(* IEC 61131-3 sources: kauha-loader-autonomy/plc/codesys/src, 6 files *)

(* ---- DUT_Types.st ---- *)
(* KAUHA safety PLC: data types.
   IEC 61131-3 Structured Text, 2nd edition subset (no methods, no references),
   so the same source compiles in CODESYS and in the matiec compiler the tests use. *)

TYPE ST_SafetyConfig :
STRUCT
    (* SafetyParams *)
    remote_timeout_s     : LREAL;
    watchdog_timeout_s   : LREAL;
    overspeed_tol        : LREAL;
    decel_ramp           : LREAL;
    ramp_reaction_s      : LREAL;
    discrepancy_tol      : LREAL;
    discrepancy_time_s   : LREAL;
    position_invalid_s   : LREAL;
    max_mute_s           : LREAL;
    auto_restart_clear_s : LREAL;
    warning_hold_s       : LREAL;
    auto_speed           : LREAL;
    teleop_speed         : LREAL;
    warning_speed        : LREAL;
    standstill           : LREAL;
    recovery_speed       : LREAL;
    side_recovery_speed  : LREAL;
    (* FieldTable: facts about the field sets loaded into the scanners *)
    t_standstill         : LREAL;
    dig_speed            : LREAL;
    dock_speed           : LREAL;
    speed_cap            : LREAL;
    auto_restart         : BOOL;     (* SR-11 automatic restart after a clearing stop *)
    band0                : LREAL;    (* speed band tops, m/s *)
    band1                : LREAL;
    band2                : LREAL;
    band3                : LREAL;
    sector0              : LREAL;    (* articulation sector boundaries, rad *)
    sector1              : LREAL;
    sector2              : LREAL;
    sector3              : LREAL;
    vprot0               : LREAL;    (* highest speed each band's protective field stops from *)
    vprot1               : LREAL;
    vprot2               : LREAL;
    vprot3               : LREAL;
    n_sectors            : INT;
    n_bands              : INT;
END_STRUCT;
END_TYPE

TYPE ST_SafetyInputs :
STRUCT
    t                : LREAL;   (* monotonic time, s *)
    mode             : INT;     (* 0 IDLE, 1 AUTO, 2 TELEOP *)
    speed_a          : LREAL;   (* drive-by-wire gateway, non-safety source, m/s *)
    speed_b          : LREAL;   (* PLC's own speed sensor, m/s *)
    articulation     : LREAL;   (* PLC's own articulation sensor, rad *)
    front_prot       : BOOL;
    front_warn       : BOOL;
    rear_prot        : BOOL;
    rear_warn        : BOOL;
    side_prot        : BOOL;
    side_contact     : BOOL;
    scanners_ok      : BOOL;
    remote_hb_age    : LREAL;
    remote_estop     : BOOL;
    reset_req        : BOOL;
    machine_estop    : BOOL;
    autonomy_cmd_age : LREAL;
    dig_req          : BOOL;
    dock_req         : BOOL;
    in_operating_area : BOOL;
    in_dig_zone      : BOOL;
    in_dock_zone     : BOOL;
    truck_door_open  : BOOL;
    boom_raised      : BOOL;
    front_side       : BOOL;
    under_near       : BOOL;
    under_far        : BOOL;
    under_mid        : BOOL;
    position_valid   : BOOL;
END_STRUCT;
END_TYPE

TYPE ST_SafetyOutputs :
STRUCT
    state            : INT;     (* 0 RUN, 1 WARNING, 2 PROTECTIVE_STOP, 3 EMERGENCY_STOP *)
    cause            : WORD;    (* latched causes, bit mask as in kauha/safety/core.py *)
    speed_limit      : LREAL;
    field_set        : INT;
    brake_release    : BOOL;    (* FALSE: drive power cut, motors short-braked (hardwired) *)
    implement_enable : BOOL;    (* FALSE: actuator power cut (hardwired) *)
    reset_pending    : BOOL;
    dock_blocked     : BOOL;
    fs_direction     : INT;
    fs_v_protected   : LREAL;
    recovery         : WORD;    (* fields in SR-12 recovery *)
    ev_stop          : BOOL;    (* a stop event was logged this cycle *)
    ev_recovery      : BOOL;
    ev_reset         : BOOL;
END_STRUCT;
END_TYPE

(* Eight payload bytes. A struct, not a bare array type, so it can be passed to
   functions by value in every IEC compiler (matiec mis-handles bare array types). *)
TYPE ST_Payload :
STRUCT
    b : ARRAY [0..7] OF BYTE;
END_STRUCT;
END_TYPE

TYPE ST_Frame :
STRUCT
    id   : DWORD;                    (* 29-bit J1939 identifier *)
    data : ST_Payload;
END_STRUCT;
END_TYPE

(* ---- GVL_Config.st ---- *)
(* KAUHA safety configuration lists, one per profile. Select one in PRG_Safety. *)

(* Generated by kauha.scale.profile for profile 'full'. Do not edit by hand. *)
VAR_GLOBAL CONSTANT
    CFG_FULL : ST_SafetyConfig := (
        remote_timeout_s := 0.5,
        watchdog_timeout_s := 0.2,
        overspeed_tol := 0.2,
        decel_ramp := 0.8,
        ramp_reaction_s := 0.3,
        discrepancy_tol := 0.3,
        discrepancy_time_s := 0.2,
        position_invalid_s := 2,
        max_mute_s := 25,
        auto_restart_clear_s := 3,
        warning_hold_s := 2,
        auto_speed := 3,
        teleop_speed := 3,
        warning_speed := 1,
        standstill := 0.05,
        recovery_speed := 0.5,
        side_recovery_speed := 0.3,
        t_standstill := 0.1,
        dig_speed := 1,
        dock_speed := 0.6,
        speed_cap := 2.97018412,
        auto_restart := TRUE,
        band0 := 0.5,
        band1 := 1.5,
        band2 := 2.5,
        band3 := 3,
        sector0 := -0.3,
        sector1 := -0.1,
        sector2 := 0.1,
        sector3 := 0.3,
        vprot0 := 0.794930202,
        vprot1 := 1.5,
        vprot2 := 2.5,
        vprot3 := 3.17018412,
        n_sectors := 5,
        n_bands := 4
    );
END_VAR

(* Generated by kauha.scale.profile for profile 'scale8_nanoscan3'. Do not edit by hand. *)
VAR_GLOBAL CONSTANT
    CFG_SCALE8_NANOSCAN3 : ST_SafetyConfig := (
        remote_timeout_s := 0.5,
        watchdog_timeout_s := 0.2,
        overspeed_tol := 0.0707106781,
        decel_ramp := 0.8,
        ramp_reaction_s := 0.1,
        discrepancy_tol := 0.106066017,
        discrepancy_time_s := 0.2,
        position_invalid_s := 2,
        max_mute_s := 8.83883476,
        auto_restart_clear_s := 1.06066017,
        warning_hold_s := 0.707106781,
        auto_speed := 1.06066017,
        teleop_speed := 1.06066017,
        warning_speed := 0.353553391,
        standstill := 0.0176776695,
        recovery_speed := 0.176776695,
        side_recovery_speed := 0.106066017,
        t_standstill := 0.0353553391,
        dig_speed := 0.353553391,
        dock_speed := 0.212132034,
        speed_cap := 1.00147274,
        auto_restart := TRUE,
        band0 := 0.176776695,
        band1 := 0.530330086,
        band2 := 0.883883476,
        band3 := 1.06066017,
        sector0 := -0.3,
        sector1 := -0.1,
        sector2 := 0.1,
        sector3 := 0.3,
        vprot0 := 0.293061951,
        vprot1 := 0.530330086,
        vprot2 := 0.883883476,
        vprot3 := 1.07218342,
        n_sectors := 5,
        n_bands := 4
    );
END_VAR

(* Generated by kauha.scale.profile for profile 'scale8_evaluator'. Do not edit by hand. *)
VAR_GLOBAL CONSTANT
    CFG_SCALE8_EVALUATOR : ST_SafetyConfig := (
        remote_timeout_s := 0.5,
        watchdog_timeout_s := 0.2,
        overspeed_tol := 0.0707106781,
        decel_ramp := 0.8,
        ramp_reaction_s := 0.1,
        discrepancy_tol := 0.106066017,
        discrepancy_time_s := 0.2,
        position_invalid_s := 2,
        max_mute_s := 8.83883476,
        auto_restart_clear_s := 1.06066017,
        warning_hold_s := 0.707106781,
        auto_speed := 1.06066017,
        teleop_speed := 1.06066017,
        warning_speed := 0.353553391,
        standstill := 0.0176776695,
        recovery_speed := 0.176776695,
        side_recovery_speed := 0.106066017,
        t_standstill := 0.0353553391,
        dig_speed := 0.353553391,
        dock_speed := 0.212132034,
        speed_cap := 0.81813501,
        auto_restart := TRUE,
        band0 := 0.176776695,
        band1 := 0.530330086,
        band2 := 0.883883476,
        band3 := 1.06066017,
        sector0 := -0.3,
        sector1 := -0.1,
        sector2 := 0.1,
        sector3 := 0.3,
        vprot0 := 0.19593478,
        vprot1 := 0.530330086,
        vprot2 := 0.883883476,
        vprot3 := 0.888845688,
        n_sectors := 5,
        n_bands := 4
    );
END_VAR

(* ---- FUN_Helpers.st ---- *)
(* Small helpers shared by the safety POUs. FMIN/FMAX reproduce the reference
   model's Min/Max exactly (first argument on ties), so results are bit-identical. *)

FUNCTION FMIN : LREAL
VAR_INPUT
    a : LREAL;
    b : LREAL;
END_VAR
FMIN := SEL(a <= b, b, a);
END_FUNCTION

FUNCTION FMAX : LREAL
VAR_INPUT
    a : LREAL;
    b : LREAL;
END_VAR
FMAX := SEL(a >= b, b, a);
END_FUNCTION

FUNCTION HAS : BOOL
VAR_INPUT
    mask : WORD;
    bits : WORD;
END_VAR
HAS := (mask AND bits) <> 0;
END_FUNCTION

(* ---- FB_SafetyCore.st ---- *)
(* KAUHA safety PLC: one 25 ms cycle of the safety logic.

   This is a line-by-line port of kauha/safety/core.py step(), the reference that
   the z3 proofs (120 properties) and the adversarial searches run on. The test
   tests/plc/test_st_equivalence.py compiles this file with matiec and checks it
   against the reference on long random and scripted input sequences: every
   output and every memory value must match bit for bit.

   Keep it that way: change core.py first, prove it, then port the change here
   and rerun the equivalence test. Requirement tags (SR-xx) follow core.py. *)

FUNCTION_BLOCK FB_SafetyCore
VAR_INPUT
    cfg : ST_SafetyConfig;
    inp : ST_SafetyInputs;
END_VAR
VAR_OUTPUT
    out : ST_SafetyOutputs;
END_VAR
VAR
    (* memory between cycles (core.Memory) *)
    m_state      : INT := 0;
    m_latched    : WORD := 0;
    m_field_set  : INT := 0;
    m_recovery   : WORD := 0;
    m_prev_reset : BOOL := FALSE;
    m_over_on    : BOOL := FALSE;
    m_over_t0    : LREAL := 0.0;
    m_disc_on    : BOOL := FALSE;
    m_disc_t0    : LREAL := 0.0;
    m_posinv_on  : BOOL := FALSE;
    m_posinv_t0  : LREAL := 0.0;
    m_mute_on    : BOOL := FALSE;
    m_mute_t0    : LREAL := 0.0;
    m_clear_on   : BOOL := FALSE;
    m_clear_t0   : LREAL := 0.0;
    m_warn_until : LREAL := -1.0;
    m_allowed    : LREAL := 0.0;
    m_prev_limit : LREAL := 0.0;
    m_env_t0     : LREAL := -1.0E9;
    m_env_v0     : LREAL := 0.0;
    (* cycle temporaries *)
    t, v, a_v       : LREAL;
    st              : INT;
    lat, rec        : WORD;
    c               : BOOL;
    ev_stop         : BOOL;
    rising_reset    : BOOL;
    dig_ok, dock_ok : BOOL;
    muting          : BOOL;
    mute_t0, posinv_t0, disc_t0, over_t0, clear_t0 : LREAL;
    mute_timeout    : BOOL;
    dig_sel, dock_sel, still : BOOL;
    sector, band, base, moving_id : INT;
    fs_id, fs_dir   : INT;
    v_band, fs_vprot : LREAL;
    at_rest         : BOOL;
    exempt, under   : BOOL;
    active_mode, is_auto, posinv, posinv_on, disc : BOOL;
    in_zone, warn_trig, warning : BOOL;
    warn_until      : LREAL;
    spd_lim, creep, env_t0, env_v0, env_ramp, allowed : LREAL;
    dec, over, travel_set, standstill : BOOL;
    active, remaining : WORD;
    stopped_now, enter_rec, clear_on, auto_ok, do_reset, stopped : BOOL;
END_VAR
VAR CONSTANT
    RUN_ST : INT := 0;
    WARNING_ST : INT := 1;
    PROTECTIVE_STOP : INT := 2;
    EMERGENCY_STOP : INT := 3;
    MODE_IDLE : INT := 0;
    MODE_AUTO : INT := 1;
    MODE_TELEOP : INT := 2;
    FIELD_FRONT : WORD := 16#0001;
    FIELD_REAR : WORD := 16#0002;
    FIELD_SIDE : WORD := 16#0004;
    OVERSPEED : WORD := 16#0008;
    REMOTE_LINK : WORD := 16#0010;
    WATCHDOG : WORD := 16#0020;
    GEOFENCE : WORD := 16#0040;
    SPEED_DISCREPANCY : WORD := 16#0080;
    SCANNER_FAULT : WORD := 16#0100;
    MUTING_TIMEOUT : WORD := 16#0200;
    ESTOP_MACHINE : WORD := 16#0400;
    ESTOP_REMOTE : WORD := 16#0800;
    POSITION_INVALID : WORD := 16#1000;
    TRUCK_DOOR : WORD := 16#2000;
    UNDER_BUCKET : WORD := 16#4000;
    FIELD_CAUSES : WORD := 16#4007;      (* FRONT | REAR | SIDE | UNDER_BUCKET *)
    CLEARING_CAUSES : WORD := 16#6007;   (* FIELD_CAUSES | TRUCK_DOOR *)
    CYCLE_S : LREAL := 0.025;
    DIG_SET : INT := 100;
    DOCK_SET : INT := 101;
    STANDSTILL_SET : INT := 0;
END_VAR

t := inp.t;
v := inp.speed_b;
st := m_state;
lat := m_latched;
ev_stop := FALSE;
out.ev_recovery := FALSE;
out.ev_reset := FALSE;

rising_reset := inp.reset_req AND NOT m_prev_reset;

(* SR-01 emergency stops: latch. *)
c := inp.machine_estop;
IF c THEN
    IF (EMERGENCY_STOP > st) OR ((ESTOP_MACHINE AND NOT lat) <> 0) THEN ev_stop := TRUE; END_IF;
    lat := lat OR ESTOP_MACHINE;
    IF EMERGENCY_STOP > st THEN st := EMERGENCY_STOP; END_IF;
END_IF;
c := inp.remote_estop;
IF c THEN
    IF (EMERGENCY_STOP > st) OR ((ESTOP_REMOTE AND NOT lat) <> 0) THEN ev_stop := TRUE; END_IF;
    lat := lat OR ESTOP_REMOTE;
    IF EMERGENCY_STOP > st THEN st := EMERGENCY_STOP; END_IF;
END_IF;

(* Field-set selection (SR-02, SR-10, SR-14). *)
dig_ok := inp.dig_req AND inp.in_dig_zone AND (ABS(v) <= cfg.dig_speed + cfg.overspeed_tol) AND inp.position_valid;
dock_ok := inp.dock_req AND inp.in_dock_zone AND (ABS(v) <= cfg.dock_speed + cfg.overspeed_tol)
           AND inp.position_valid AND NOT inp.truck_door_open;
(* SR-14: the driver leaving the cab while the loader is docking stops it. *)
c := inp.truck_door_open AND (m_field_set = DOCK_SET) AND inp.in_dock_zone;
IF c THEN
    IF (PROTECTIVE_STOP > st) OR ((TRUCK_DOOR AND NOT lat) <> 0) THEN ev_stop := TRUE; END_IF;
    lat := lat OR TRUCK_DOOR;
    IF PROTECTIVE_STOP > st THEN st := PROTECTIVE_STOP; END_IF;
END_IF;
muting := dig_ok AND (v > -cfg.t_standstill);
mute_t0 := SEL(muting AND m_mute_on, t, m_mute_t0);
mute_timeout := muting AND (t - mute_t0 > cfg.max_mute_s);
c := mute_timeout;
IF c THEN
    IF (PROTECTIVE_STOP > st) OR ((MUTING_TIMEOUT AND NOT lat) <> 0) THEN ev_stop := TRUE; END_IF;
    lat := lat OR MUTING_TIMEOUT;
    IF PROTECTIVE_STOP > st THEN st := PROTECTIVE_STOP; END_IF;
END_IF;
dig_ok := dig_ok AND NOT mute_timeout;

(* select(): set id, direction, protected speed *)
dig_sel := dig_ok AND (v > -cfg.t_standstill);
dock_sel := NOT dig_sel AND dock_ok AND (v > -cfg.t_standstill);
still := ABS(v) < cfg.t_standstill;
a_v := ABS(v);
IF inp.articulation < cfg.sector0 THEN sector := 0;
ELSIF inp.articulation < cfg.sector1 THEN sector := 1;
ELSIF inp.articulation < cfg.sector2 THEN sector := 2;
ELSIF inp.articulation < cfg.sector3 THEN sector := 3;
ELSE sector := 4;
END_IF;
IF a_v <= cfg.band0 THEN band := 0;
ELSIF a_v <= cfg.band1 THEN band := 1;
ELSIF a_v <= cfg.band2 THEN band := 2;
ELSE band := 3;
END_IF;
base := SEL(v > 0.0, 1 + cfg.n_bands * cfg.n_sectors, 1);
moving_id := base + band * cfg.n_sectors + sector;
IF dig_sel THEN fs_id := DIG_SET;
ELSIF dock_sel THEN fs_id := DOCK_SET;
ELSIF still THEN fs_id := STANDSTILL_SET;
ELSE fs_id := moving_id;
END_IF;
IF dig_sel OR dock_sel THEN fs_dir := 1;
ELSIF still THEN fs_dir := 0;
ELSIF v > 0.0 THEN fs_dir := 1;
ELSE fs_dir := -1;
END_IF;
IF band = 0 THEN v_band := cfg.vprot0;
ELSIF band = 1 THEN v_band := cfg.vprot1;
ELSIF band = 2 THEN v_band := cfg.vprot2;
ELSE v_band := cfg.vprot3;
END_IF;
IF dig_sel THEN fs_vprot := cfg.dig_speed;
ELSIF dock_sel THEN fs_vprot := cfg.dock_speed;
ELSIF still THEN fs_vprot := cfg.t_standstill;
ELSE fs_vprot := v_band;
END_IF;

(* SR-12 recovery: after a supervisor reset in TELEOP, motion away from an occupied
   field is allowed at creep speed; motion toward it trips again. A field counts as
   clear only at standstill. *)
rec := SEL(inp.mode = MODE_TELEOP, WORD#0, m_recovery);
at_rest := ABS(v) < cfg.standstill;
IF at_rest AND NOT inp.front_prot THEN rec := rec AND NOT FIELD_FRONT; END_IF;
IF at_rest AND NOT inp.rear_prot THEN rec := rec AND NOT FIELD_REAR; END_IF;
IF at_rest AND NOT inp.side_prot THEN rec := rec AND NOT FIELD_SIDE; END_IF;
(* SR-16: someone between the front tyres and the bucket, or under the raised bucket. *)
exempt := inp.in_dig_zone OR (inp.in_dock_zone AND NOT inp.truck_door_open);
under := NOT inp.in_dig_zone AND (inp.under_near OR (NOT exempt AND (inp.under_mid OR (inp.boom_raised AND inp.under_far))));
IF at_rest AND NOT under THEN rec := rec AND NOT UNDER_BUCKET; END_IF;

c := HAS(rec, FIELD_SIDE) AND inp.side_contact AND NOT exempt;
IF c THEN
    IF (PROTECTIVE_STOP > st) OR ((FIELD_SIDE AND NOT lat) <> 0) THEN ev_stop := TRUE; END_IF;
    lat := lat OR FIELD_SIDE;
    IF PROTECTIVE_STOP > st THEN st := PROTECTIVE_STOP; END_IF;
END_IF;
c := HAS(rec, UNDER_BUCKET) AND (v > cfg.standstill);
IF c THEN
    IF (PROTECTIVE_STOP > st) OR ((UNDER_BUCKET AND NOT lat) <> 0) THEN ev_stop := TRUE; END_IF;
    lat := lat OR UNDER_BUCKET;
    IF PROTECTIVE_STOP > st THEN st := PROTECTIVE_STOP; END_IF;
END_IF;
c := HAS(rec, FIELD_FRONT) AND (v > cfg.standstill);
IF c THEN
    IF (PROTECTIVE_STOP > st) OR ((FIELD_FRONT AND NOT lat) <> 0) THEN ev_stop := TRUE; END_IF;
    lat := lat OR FIELD_FRONT;
    IF PROTECTIVE_STOP > st THEN st := PROTECTIVE_STOP; END_IF;
END_IF;
c := HAS(rec, FIELD_REAR) AND (v < -cfg.standstill);
IF c THEN
    IF (PROTECTIVE_STOP > st) OR ((FIELD_REAR AND NOT lat) <> 0) THEN ev_stop := TRUE; END_IF;
    lat := lat OR FIELD_REAR;
    IF PROTECTIVE_STOP > st THEN st := PROTECTIVE_STOP; END_IF;
END_IF;

(* SR-02 protective fields. The scanners evaluate the selected set. *)
c := inp.front_prot AND (fs_dir >= 0) AND NOT HAS(rec, FIELD_FRONT);
IF c THEN
    IF (PROTECTIVE_STOP > st) OR ((FIELD_FRONT AND NOT lat) <> 0) THEN ev_stop := TRUE; END_IF;
    lat := lat OR FIELD_FRONT;
    IF PROTECTIVE_STOP > st THEN st := PROTECTIVE_STOP; END_IF;
END_IF;
c := inp.rear_prot AND ((fs_dir <= 0) OR (ABS(v) < cfg.standstill)) AND NOT HAS(rec, FIELD_REAR);
IF c THEN
    IF (PROTECTIVE_STOP > st) OR ((FIELD_REAR AND NOT lat) <> 0) THEN ev_stop := TRUE; END_IF;
    lat := lat OR FIELD_REAR;
    IF PROTECTIVE_STOP > st THEN st := PROTECTIVE_STOP; END_IF;
END_IF;
c := inp.side_prot AND (ABS(v) > cfg.standstill) AND NOT HAS(rec, FIELD_SIDE);
IF c THEN
    IF (PROTECTIVE_STOP > st) OR ((FIELD_SIDE AND NOT lat) <> 0) THEN ev_stop := TRUE; END_IF;
    lat := lat OR FIELD_SIDE;
    IF PROTECTIVE_STOP > st THEN st := PROTECTIVE_STOP; END_IF;
END_IF;
c := NOT inp.scanners_ok;
IF c THEN
    IF (PROTECTIVE_STOP > st) OR ((SCANNER_FAULT AND NOT lat) <> 0) THEN ev_stop := TRUE; END_IF;
    lat := lat OR SCANNER_FAULT;
    IF PROTECTIVE_STOP > st THEN st := PROTECTIVE_STOP; END_IF;
END_IF;
(* SR-16: a person under the raised bucket stops travel and holds the boom. *)
c := under AND NOT HAS(rec, UNDER_BUCKET);
IF c THEN
    IF (PROTECTIVE_STOP > st) OR ((UNDER_BUCKET AND NOT lat) <> 0) THEN ev_stop := TRUE; END_IF;
    lat := lat OR UNDER_BUCKET;
    IF PROTECTIVE_STOP > st THEN st := PROTECTIVE_STOP; END_IF;
END_IF;
(* Reversing: someone stepping in beside the front frame heads for the gap between
   the front tyres and the bucket's back edge. *)
c := inp.front_side AND (v < -cfg.standstill) AND NOT exempt AND NOT HAS(rec, FIELD_SIDE);
IF c THEN
    IF (PROTECTIVE_STOP > st) OR ((FIELD_SIDE AND NOT lat) <> 0) THEN ev_stop := TRUE; END_IF;
    lat := lat OR FIELD_SIDE;
    IF PROTECTIVE_STOP > st THEN st := PROTECTIVE_STOP; END_IF;
END_IF;

(* SR-05 remote supervision link, SR-06 autonomy watchdog. *)
active_mode := (inp.mode = MODE_AUTO) OR (inp.mode = MODE_TELEOP);
c := active_mode AND (inp.remote_hb_age > cfg.remote_timeout_s);
IF c THEN
    IF (PROTECTIVE_STOP > st) OR ((REMOTE_LINK AND NOT lat) <> 0) THEN ev_stop := TRUE; END_IF;
    lat := lat OR REMOTE_LINK;
    IF PROTECTIVE_STOP > st THEN st := PROTECTIVE_STOP; END_IF;
END_IF;
c := active_mode AND (inp.autonomy_cmd_age > cfg.watchdog_timeout_s);
IF c THEN
    IF (PROTECTIVE_STOP > st) OR ((WATCHDOG AND NOT lat) <> 0) THEN ev_stop := TRUE; END_IF;
    lat := lat OR WATCHDOG;
    IF PROTECTIVE_STOP > st THEN st := PROTECTIVE_STOP; END_IF;
END_IF;

(* SR-07 geofence; an invalid position is tolerated briefly. *)
is_auto := inp.mode = MODE_AUTO;
posinv := is_auto AND NOT inp.position_valid;
posinv_t0 := SEL(posinv AND NOT m_posinv_on, m_posinv_t0, t);
posinv_on := SEL(is_auto, m_posinv_on, NOT inp.position_valid);
c := posinv AND (t - posinv_t0 > cfg.position_invalid_s);
IF c THEN
    IF (PROTECTIVE_STOP > st) OR ((POSITION_INVALID AND NOT lat) <> 0) THEN ev_stop := TRUE; END_IF;
    lat := lat OR POSITION_INVALID;
    IF PROTECTIVE_STOP > st THEN st := PROTECTIVE_STOP; END_IF;
END_IF;
c := is_auto AND inp.position_valid AND NOT inp.in_operating_area;
IF c THEN
    IF (PROTECTIVE_STOP > st) OR ((GEOFENCE AND NOT lat) <> 0) THEN ev_stop := TRUE; END_IF;
    lat := lat OR GEOFENCE;
    IF PROTECTIVE_STOP > st THEN st := PROTECTIVE_STOP; END_IF;
END_IF;

(* SR-08 two-channel speed plausibility. *)
disc := ABS(inp.speed_a - inp.speed_b) > cfg.discrepancy_tol;
disc_t0 := SEL(disc AND NOT m_disc_on, m_disc_t0, t);
c := disc AND (t - disc_t0 > cfg.discrepancy_time_s);
IF c THEN
    IF (PROTECTIVE_STOP > st) OR ((SPEED_DISCREPANCY AND NOT lat) <> 0) THEN ev_stop := TRUE; END_IF;
    lat := lat OR SPEED_DISCREPANCY;
    IF PROTECTIVE_STOP > st THEN st := PROTECTIVE_STOP; END_IF;
END_IF;

(* SR-03 warning field -> speed limit (non-latching), not inside the dig and dock zones. *)
in_zone := inp.in_dig_zone OR inp.in_dock_zone;
warn_trig := NOT in_zone AND ((inp.front_warn AND (fs_dir >= 0)) OR (inp.rear_warn AND (fs_dir <= 0)));
warn_until := SEL(warn_trig, m_warn_until, t + cfg.warning_hold_s);
warning := t < warn_until;

(* SR-04 speed limit and overspeed monitoring. *)
IF is_auto THEN
    spd_lim := FMIN(cfg.auto_speed, cfg.speed_cap);
ELSIF inp.mode = MODE_TELEOP THEN
    spd_lim := FMIN(cfg.teleop_speed, cfg.speed_cap);
ELSE
    spd_lim := 0.0;
END_IF;
IF warning THEN spd_lim := FMIN(spd_lim, cfg.warning_speed); END_IF;
creep := SEL(HAS(rec, FIELD_SIDE), cfg.recovery_speed, cfg.side_recovery_speed);
IF rec <> 0 THEN spd_lim := FMIN(spd_lim, creep); END_IF;
IF fs_id = DIG_SET THEN
    spd_lim := FMIN(spd_lim, cfg.dig_speed);
ELSIF fs_id = DOCK_SET THEN
    spd_lim := FMIN(spd_lim, cfg.dock_speed);
END_IF;
(* The monitored envelope follows a limit increase at once; after a decrease it holds
   the current speed for the reaction time, then ramps down (SS1-r style). *)
dec := spd_lim < m_prev_limit - 1.0E-9;
env_t0 := SEL(dec, m_env_t0, t);
env_v0 := SEL(dec, m_env_v0, FMIN(m_allowed, ABS(v)));
env_ramp := env_v0 - cfg.decel_ramp * FMAX(0.0, t - env_t0 - cfg.ramp_reaction_s);
allowed := FMAX(spd_lim, env_ramp);
over := ABS(v) > allowed + cfg.overspeed_tol;
over_t0 := SEL(over AND NOT m_over_on, m_over_t0, t);
c := over AND (t - over_t0 >= CYCLE_S);
IF c THEN
    IF (PROTECTIVE_STOP > st) OR ((OVERSPEED AND NOT lat) <> 0) THEN ev_stop := TRUE; END_IF;
    lat := lat OR OVERSPEED;
    IF PROTECTIVE_STOP > st THEN st := PROTECTIVE_STOP; END_IF;
END_IF;
(* Never travel faster than the selected protective field can stop from. *)
travel_set := (fs_dir <> 0) AND (fs_id <> DIG_SET) AND (fs_id <> DOCK_SET);
c := travel_set AND (ABS(v) > fs_vprot);
IF c THEN
    IF (PROTECTIVE_STOP > st) OR ((OVERSPEED AND NOT lat) <> 0) THEN ev_stop := TRUE; END_IF;
    lat := lat OR OVERSPEED;
    IF PROTECTIVE_STOP > st THEN st := PROTECTIVE_STOP; END_IF;
END_IF;

(* Reset handling (SR-09, SR-11, SR-12). *)
standstill := ABS(v) < cfg.standstill;
active := 0;
IF inp.machine_estop THEN active := active OR ESTOP_MACHINE; END_IF;
IF inp.remote_estop THEN active := active OR ESTOP_REMOTE; END_IF;
IF inp.front_prot THEN active := active OR FIELD_FRONT; END_IF;
IF inp.rear_prot THEN active := active OR FIELD_REAR; END_IF;
IF inp.side_prot THEN active := active OR FIELD_SIDE; END_IF;
IF NOT inp.scanners_ok THEN active := active OR SCANNER_FAULT; END_IF;
IF (inp.mode <> MODE_IDLE) AND (inp.remote_hb_age > cfg.remote_timeout_s) THEN active := active OR REMOTE_LINK; END_IF;
IF (inp.mode <> MODE_IDLE) AND (inp.autonomy_cmd_age > cfg.watchdog_timeout_s) THEN active := active OR WATCHDOG; END_IF;
IF is_auto AND inp.position_valid AND NOT inp.in_operating_area THEN active := active OR GEOFENCE; END_IF;
IF ABS(inp.speed_a - inp.speed_b) > cfg.discrepancy_tol THEN active := active OR SPEED_DISCREPANCY; END_IF;
IF is_auto AND NOT inp.position_valid THEN active := active OR POSITION_INVALID; END_IF;
IF inp.truck_door_open AND inp.in_dock_zone THEN active := active OR TRUCK_DOOR; END_IF;
IF under THEN active := active OR UNDER_BUCKET; END_IF;
(* Muting past its limit blocks reset while the dig request continues. *)
IF mute_timeout THEN active := active OR MUTING_TIMEOUT; END_IF;
(* A cause latched in this very cycle cannot be reset in the same cycle. *)
stopped_now := (st >= PROTECTIVE_STOP) AND NOT ((lat AND NOT m_latched) <> 0);
remaining := lat AND active;
enter_rec := stopped_now AND rising_reset AND (inp.mode = MODE_TELEOP) AND (st = PROTECTIVE_STOP)
             AND (remaining <> 0) AND ((remaining AND NOT FIELD_CAUSES) = 0)
             AND NOT (HAS(remaining, FIELD_SIDE) AND inp.side_contact AND NOT exempt);
(* Fields already in recovery stay in it. *)
IF enter_rec THEN rec := rec OR remaining; END_IF;
out.ev_recovery := enter_rec;
IF enter_rec THEN remaining := 0; END_IF;
clear_t0 := SEL(stopped_now AND (remaining = 0) AND NOT m_clear_on, m_clear_t0, t);
clear_on := SEL(stopped_now, m_clear_on, remaining = 0);
IF cfg.auto_restart THEN
    auto_ok := (st = PROTECTIVE_STOP) AND ((lat AND NOT CLEARING_CAUSES) = 0) AND clear_on
               AND (t - clear_t0 >= cfg.auto_restart_clear_s) AND NOT warning;
ELSE
    auto_ok := FALSE;
END_IF;
do_reset := stopped_now AND standstill AND (remaining = 0) AND (rising_reset OR auto_ok);
out.ev_reset := do_reset;
IF do_reset THEN
    st := RUN_ST;
    lat := 0;
    clear_on := FALSE;
END_IF;
IF st < PROTECTIVE_STOP THEN
    st := SEL(warning, RUN_ST, WARNING_ST);
END_IF;

stopped := st >= PROTECTIVE_STOP;
m_state := st;
m_latched := lat;
m_field_set := fs_id;
m_recovery := rec;
m_prev_reset := inp.reset_req;
m_over_on := over;
m_over_t0 := over_t0;
m_disc_on := disc;
m_disc_t0 := disc_t0;
m_posinv_on := posinv_on;
m_posinv_t0 := posinv_t0;
m_mute_on := muting;
m_mute_t0 := mute_t0;
m_clear_on := clear_on;
m_clear_t0 := clear_t0;
m_warn_until := warn_until;
m_allowed := allowed;
m_prev_limit := spd_lim;
m_env_t0 := env_t0;
m_env_v0 := env_v0;

(* The recovery creep limit applies from the cycle recovery starts. *)
creep := SEL(HAS(rec, FIELD_SIDE), cfg.recovery_speed, cfg.side_recovery_speed);
IF rec <> 0 THEN spd_lim := FMIN(spd_lim, creep); END_IF;
out.state := st;
out.cause := lat;
out.speed_limit := SEL(stopped, spd_lim, 0.0);
out.field_set := fs_id;
out.brake_release := NOT stopped;
(* SR-12: no boom/bucket motion while recovering from an occupied field. *)
out.implement_enable := NOT stopped AND (rec = 0);
out.reset_pending := stopped AND ((lat AND active) = 0);
out.dock_blocked := inp.truck_door_open;
out.fs_direction := fs_dir;
out.fs_v_protected := fs_vprot;
out.recovery := rec;
out.ev_stop := ev_stop;
END_FUNCTION_BLOCK

(* ---- FB_SafetyNode.st ---- *)
(* KAUHA safety PLC, testbed node: everything between the CAN driver and the
   safety core, in plain IEC 61131-3 so it is tested with the core.

   Each 25 ms cycle PRG_Main (CODESYS-specific CAN driver calls) hands this block
   the frames received since the last cycle and the GPIO inputs. It checks every
   frame end to end (CRC, alive counter, freshness), builds the core's inputs,
   runs FB_SafetyCore, and returns the SafetyStatus frame and the hardwired outputs.

   Fail-safe defaults: a frame that is missing, stale or corrupt never makes the
   machine run; see the comment at each input. *)

TYPE ST_RxBatch :
STRUCT
    n : INT;                               (* frames valid in f[0..n-1] *)
    f : ARRAY [0..31] OF ST_Frame;
END_STRUCT;
END_TYPE

TYPE ST_ScannerIO :
STRUCT
    (* Rated scanner option (SICK nanoScan3 I/O or similar), wired to PLC inputs.
       OSSD-type signals are TRUE when the field is CLEAR. *)
    front_ossd_clear : BOOL;
    rear_ossd_clear  : BOOL;
    front_warn_clear : BOOL;
    rear_warn_clear  : BOOL;
    side_clear       : BOOL;
    under_clear      : BOOL;    (* under_near and under_mid share one output on the testbed *)
    scanners_ready   : BOOL;    (* scanner "device ready / no fault" outputs, both scanners *)
END_STRUCT;
END_TYPE

FUNCTION_BLOCK FB_SafetyNode
VAR_INPUT
    cfg            : ST_SafetyConfig;
    t              : LREAL;          (* s, monotonic *)
    rx             : ST_RxBatch;
    estop_chain_ok : BOOL;           (* machine e-stop chain closed: safety relay K1 output state *)
    use_scanner_io : BOOL;           (* TRUE: rated scanner outputs on GPIO; FALSE: ScannerStatus frames *)
    scanner_io     : ST_ScannerIO;
END_VAR
VAR_OUTPUT
    out              : ST_SafetyOutputs;
    drive_enable     : BOOL;         (* relay K-DRIVE: motor power and dynamic-brake changeover *)
    implement_enable : BOOL;         (* relay K-IMPL: actuator power *)
    field_set_code   : BYTE;         (* to the rated scanners' static control inputs *)
    tx_id            : DWORD;
    tx               : ST_Payload;   (* SafetyStatus, protected *)
    inputs           : ST_SafetyInputs;   (* what the core saw this cycle, for diagnostics *)
    sensor_fault     : BOOL;
    scanner_fault    : BOOL;
END_VAR
VAR
    core : FB_SafetyCore;
    rxDrive, rxRemote, rxMs1, rxSensors, rxScanner, rxZone : FB_E2ERx;
    k : INT;
    id : DWORD;
    pgn : DWORD;
    sa : DWORD;
    d : ST_Payload;
    (* last accepted values; start in the safe state *)
    mode_req : INT := 0;
    remote_estop : BOOL := TRUE;
    reset_req : BOOL := FALSE;
    dig_req, dock_req : BOOL := FALSE;
    speed_a : LREAL := 0.0;
    speed_b : LREAL := 0.0;
    articulation : LREAL := 0.0;
    boom_raised : BOOL := TRUE;
    sensor_ok : BOOL := FALSE;
    sc_bits : ST_Payload;
    sc_set : INT := -1;
    zone : ST_Payload;
    hist : ARRAY [0..3] OF INT := [-2, -2, -2, -2];
    set_ok : BOOL;
    counter : INT := 0;
    ok : BOOL;
END_VAR

FOR k := 0 TO rx.n - 1 DO
    id := rx.f[k].id;
    d := rx.f[k].data;
    pgn := SHR(id, 8) AND 16#3FFFF;
    sa := id AND 16#FF;
    IF (pgn = 16#FF40) AND (sa = 16#82) THEN                 (* RemoteHeartbeat *)
        rxRemote(data_id := 16#40, timeout_s := cfg.remote_timeout_s, new_frame := TRUE, data := d, t := t);
        IF rxRemote.accepted THEN
            remote_estop := GET_BIT(d, 0);
            reset_req := GET_BIT(d, 1);
            mode_req := GET_U4(d, 4);
        END_IF;
    ELSIF (pgn = 16#FF10) AND (sa = 16#80) THEN              (* DriveCmd *)
        rxDrive(data_id := 16#10, timeout_s := cfg.watchdog_timeout_s, new_frame := TRUE, data := d, t := t);
        IF rxDrive.accepted THEN
            dig_req := GET_BIT(d, 37);
            dock_req := GET_BIT(d, 38);
        END_IF;
    ELSIF (pgn = 16#FF30) AND (sa = 16#83) THEN              (* MachineState1 *)
        rxMs1(data_id := 16#30, timeout_s := 0.1, new_frame := TRUE, data := d, t := t);
        IF rxMs1.accepted THEN speed_a := GET_S16(d, 0, 0.001); END_IF;
    ELSIF (pgn = 16#FF50) AND (sa = 16#84) THEN              (* SafeSensors *)
        rxSensors(data_id := 16#50, timeout_s := 0.1, new_frame := TRUE, data := d, t := t);
        IF rxSensors.accepted THEN
            speed_b := GET_S16(d, 0, 0.001);
            articulation := GET_S16(d, 2, 0.0001);
            boom_raised := GET_BIT(d, 52);
            sensor_ok := GET_BIT(d, 53);
        END_IF;
    ELSIF (pgn = 16#FF51) AND (sa = 16#85) THEN              (* ScannerStatus *)
        rxScanner(data_id := 16#51, timeout_s := 0.1, new_frame := TRUE, data := d, t := t);
        IF rxScanner.accepted THEN
            sc_bits := d;
            sc_set := BYTE_TO_INT(d.b[2]);
        END_IF;
    ELSIF (pgn = 16#FF52) AND (sa = 16#86) THEN              (* ZoneStatus *)
        rxZone(data_id := 16#52, timeout_s := 0.5, new_frame := TRUE, data := d, t := t);
        IF rxZone.accepted THEN zone := d; END_IF;
    END_IF;
END_FOR;
(* freshness and age at this cycle's time *)
rxRemote(new_frame := FALSE, t := t);
rxDrive(new_frame := FALSE, t := t);
rxMs1(new_frame := FALSE, t := t);
rxSensors(new_frame := FALSE, t := t);
rxScanner(new_frame := FALSE, t := t);
rxZone(new_frame := FALSE, t := t);

inputs.t := t;
inputs.mode := mode_req;
(* SR-05/SR-06 run on the ages; before the first frame the age is 1E9 s. *)
inputs.remote_hb_age := rxRemote.age;
inputs.autonomy_cmd_age := rxDrive.age;
(* Stale remote: keep the e-stop state last received; the link timeout stops the machine. *)
inputs.remote_estop := remote_estop;
inputs.reset_req := reset_req AND rxRemote.fresh;
inputs.dig_req := dig_req AND rxDrive.fresh;
inputs.dock_req := dock_req AND rxDrive.fresh;
inputs.machine_estop := NOT estop_chain_ok;
(* SR-08: a silent gateway reads as a large speed, so the discrepancy check stops the machine. *)
IF rxMs1.fresh THEN inputs.speed_a := speed_a; ELSE inputs.speed_a := 1000.0; END_IF;
(* The PLC's own sensors: if stale or reporting a fault, the core sees a sensor/scanner
   fault (cause SCANNER_FAULT) and the last speed is held. *)
sensor_fault := NOT (rxSensors.fresh AND sensor_ok);
inputs.speed_b := speed_b;
inputs.articulation := articulation;
inputs.boom_raised := boom_raised OR sensor_fault;
(* Field inputs *)
IF use_scanner_io THEN
    inputs.front_prot := NOT scanner_io.front_ossd_clear;
    inputs.rear_prot := NOT scanner_io.rear_ossd_clear;
    inputs.front_warn := NOT scanner_io.front_warn_clear;
    inputs.rear_warn := NOT scanner_io.rear_warn_clear;
    inputs.side_prot := NOT scanner_io.side_clear;
    inputs.side_contact := NOT scanner_io.side_clear;
    inputs.front_side := NOT scanner_io.side_clear;
    inputs.under_near := NOT scanner_io.under_clear;
    inputs.under_mid := NOT scanner_io.under_clear;
    inputs.under_far := FALSE;
    scanner_fault := NOT scanner_io.scanners_ready;
ELSE
    (* The evaluator must be evaluating a set the PLC selected in the last four cycles. *)
    set_ok := (sc_set = hist[0]) OR (sc_set = hist[1]) OR (sc_set = hist[2]) OR (sc_set = hist[3]);
    scanner_fault := NOT (rxScanner.fresh AND GET_BIT(sc_bits, 10) AND set_ok);
    IF scanner_fault THEN
        (* every field reads occupied *)
        inputs.front_prot := TRUE; inputs.rear_prot := TRUE; inputs.front_warn := TRUE; inputs.rear_warn := TRUE;
        inputs.side_prot := TRUE; inputs.side_contact := TRUE; inputs.front_side := TRUE;
        inputs.under_near := TRUE; inputs.under_mid := TRUE; inputs.under_far := TRUE;
    ELSE
        inputs.front_prot := GET_BIT(sc_bits, 0);
        inputs.front_warn := GET_BIT(sc_bits, 1);
        inputs.rear_prot := GET_BIT(sc_bits, 2);
        inputs.rear_warn := GET_BIT(sc_bits, 3);
        inputs.side_prot := GET_BIT(sc_bits, 4);
        inputs.side_contact := GET_BIT(sc_bits, 5);
        inputs.front_side := GET_BIT(sc_bits, 6);
        inputs.under_near := GET_BIT(sc_bits, 7);
        inputs.under_mid := GET_BIT(sc_bits, 8);
        inputs.under_far := GET_BIT(sc_bits, 9);
    END_IF;
END_IF;
inputs.scanners_ok := NOT scanner_fault AND NOT sensor_fault;
(* Zones: stale means position invalid and outside every zone. *)
IF rxZone.fresh THEN
    inputs.in_operating_area := GET_BIT(zone, 0);
    inputs.in_dig_zone := GET_BIT(zone, 1);
    inputs.in_dock_zone := GET_BIT(zone, 2);
    inputs.position_valid := GET_BIT(zone, 3);
    inputs.truck_door_open := GET_BIT(zone, 4);
ELSE
    inputs.in_operating_area := FALSE;
    inputs.in_dig_zone := FALSE;
    inputs.in_dock_zone := FALSE;
    inputs.position_valid := FALSE;
    inputs.truck_door_open := TRUE;
END_IF;

core(cfg := cfg, inp := inputs);
out := core.out;

hist[3] := hist[2];
hist[2] := hist[1];
hist[1] := hist[0];
hist[0] := out.field_set;

drive_enable := out.brake_release;
implement_enable := out.implement_enable;
field_set_code := INT_TO_BYTE(out.field_set);
counter := (counter + 1) MOD 16;
tx_id := 16#08FF2081;
ok := ENCODE_SAFETY_STATUS(out, counter, 16#20, tx);
END_FUNCTION_BLOCK

(* ---- FUN_Can.st ---- *)
(* KAUHA machine bus in the safety PLC: CRC-8 (SAE J1850), end-to-end receiver,
   signal packing. Port of kauha/can/e2e.py and the frame layouts in
   hardware/can/kauha_machine.dbc (little-endian, Intel byte order).
   tests/plc/test_st_equivalence.py checks these against the Python codec. *)

FUNCTION CRC8_J1850 : BYTE
VAR_INPUT
    data_id : BYTE;
    data    : ST_Payload;   (* CRC over data_id then bytes 0..6 *)
END_VAR
VAR
    crc : BYTE;
    i, k : INT;
    nb : BYTE;
END_VAR
crc := 16#FF;
FOR i := -1 TO 6 DO
    IF i < 0 THEN nb := data_id; ELSE nb := data.b[i]; END_IF;
    crc := crc XOR nb;
    FOR k := 1 TO 8 DO
        IF (crc AND 16#80) <> 0 THEN
            crc := SHL(crc, 1) XOR 16#1D;
        ELSE
            crc := SHL(crc, 1);
        END_IF;
    END_FOR;
END_FOR;
CRC8_J1850 := crc XOR 16#FF;
END_FUNCTION

FUNCTION E2E_PROTECT : BOOL   (* writes counter and CRC into data; always TRUE *)
VAR_INPUT
    data_id : BYTE;
    counter : INT;
END_VAR
VAR_IN_OUT
    data : ST_Payload;
END_VAR
data.b[6] := (data.b[6] AND 16#F0) OR (INT_TO_BYTE(counter) AND 16#0F);
data.b[7] := CRC8_J1850(data_id, data);
E2E_PROTECT := TRUE;
END_FUNCTION

(* E2E receiver. status: 0 OK, 1 OK_SOME_LOST, 2 REPEATED, 3 WRONG_SEQUENCE, 4 CRC_ERROR.
   Call with new_frame := TRUE once per received frame; fresh is evaluated every call. *)
FUNCTION_BLOCK FB_E2ERx
VAR_INPUT
    data_id   : BYTE;
    timeout_s : LREAL;
    max_delta : INT := 2;
    new_frame : BOOL;
    data      : ST_Payload;
    t         : LREAL;
END_VAR
VAR_OUTPUT
    status : INT;
    accepted : BOOL;    (* this frame passed: OK or OK_SOME_LOST *)
    fresh  : BOOL;
    age    : LREAL;     (* seconds since the last accepted frame (1E9 before the first) *)
END_VAR
VAR
    last_counter : INT := -1;
    last_ok_time : LREAL := -1.0E9;
    have_ok : BOOL := FALSE;
    ctr, delta : INT;
END_VAR
accepted := FALSE;
IF new_frame THEN
    IF CRC8_J1850(data_id, data) <> data.b[7] THEN
        status := 4;
    ELSE
        ctr := BYTE_TO_INT(data.b[6] AND 16#0F);
        IF last_counter < 0 THEN
            status := 0;
            last_counter := ctr;
        ELSE
            delta := (ctr - last_counter + 16) MOD 16;
            IF delta = 0 THEN
                status := 2;
            ELSE
                IF delta > max_delta THEN status := 3;
                ELSIF delta = 1 THEN status := 0;
                ELSE status := 1;
                END_IF;
                last_counter := ctr;
            END_IF;
        END_IF;
        IF status <= 1 THEN
            accepted := TRUE;
            last_ok_time := t;
            have_ok := TRUE;
        END_IF;
    END_IF;
END_IF;
fresh := have_ok AND (t - last_ok_time <= timeout_s);
IF have_ok THEN age := t - last_ok_time; ELSE age := 1.0E9; END_IF;
END_FUNCTION_BLOCK

(* Signal access, Intel byte order. start_byte is the signal's start bit / 8. *)
FUNCTION GET_S16 : LREAL   (* signed 16 bit times factor *)
VAR_INPUT
    data : ST_Payload;
    start_byte : INT;
    factor : LREAL;
END_VAR
VAR
    raw : DINT;
END_VAR
raw := BYTE_TO_DINT(data.b[start_byte]) + 256 * BYTE_TO_DINT(data.b[start_byte + 1]);
IF raw >= 32768 THEN raw := raw - 65536; END_IF;
GET_S16 := DINT_TO_LREAL(raw) * factor;
END_FUNCTION

FUNCTION GET_U16 : DINT
VAR_INPUT
    data : ST_Payload;
    start_byte : INT;
END_VAR
GET_U16 := BYTE_TO_DINT(data.b[start_byte]) + 256 * BYTE_TO_DINT(data.b[start_byte + 1]);
END_FUNCTION

FUNCTION GET_BIT : BOOL
VAR_INPUT
    data : ST_Payload;
    bit : INT;            (* DBC start bit *)
END_VAR
GET_BIT := (SHR(data.b[bit / 8], bit MOD 8) AND 16#01) <> 0;
END_FUNCTION

FUNCTION GET_U4 : INT
VAR_INPUT
    data : ST_Payload;
    bit : INT;            (* DBC start bit, nibble aligned *)
END_VAR
GET_U4 := BYTE_TO_INT(SHR(data.b[bit / 8], bit MOD 8) AND 16#0F);
END_FUNCTION

FUNCTION PUT_U16 : BOOL
VAR_INPUT
    value : DINT;         (* 0..65535 *)
    start_byte : INT;
END_VAR
VAR_IN_OUT
    data : ST_Payload;
END_VAR
data.b[start_byte] := DINT_TO_BYTE(value MOD 256);
data.b[start_byte + 1] := DINT_TO_BYTE(value / 256);
PUT_U16 := TRUE;
END_FUNCTION

(* SafetyStatus frame (PLC -> gateway, autonomy, remote). Payload as the DBC:
   State 0|4, ResetPending 4|1, DockBlocked 5|1, ActiveFieldSet 8|8, Cause 16|16,
   SpeedLimit 32|16 (0.001 m/s), AliveCounter 48|4, Crc 56|8. *)
FUNCTION ENCODE_SAFETY_STATUS : BOOL
VAR_INPUT
    o : ST_SafetyOutputs;
    counter : INT;
    data_id : BYTE;
END_VAR
VAR_IN_OUT
    data : ST_Payload;
END_VAR
VAR
    i : INT;
    lim : DINT;
    ok : BOOL;
END_VAR
FOR i := 0 TO 7 DO data.b[i] := 0; END_FOR;
data.b[0] := INT_TO_BYTE(o.state) AND 16#0F;
IF o.reset_pending THEN data.b[0] := data.b[0] OR 16#10; END_IF;
IF o.dock_blocked THEN data.b[0] := data.b[0] OR 16#20; END_IF;
data.b[1] := INT_TO_BYTE(o.field_set);
ok := PUT_U16(WORD_TO_DINT(o.cause), 2, data);
lim := LREAL_TO_DINT(o.speed_limit * 1000.0);
IF lim < 0 THEN lim := 0; END_IF;
IF lim > 6000 THEN lim := 6000; END_IF;
ok := PUT_U16(lim, 4, data);
ok := E2E_PROTECT(data_id, counter, data);
ENCODE_SAFETY_STATUS := TRUE;
END_FUNCTION
